(* CODESYS project DemoLib.library
   Title: DemoLib
   Author: TwinCAT Explorer
   Company: Demo
   Version: 1.0.0.0
   Placeholder: DemoLib

Project tree, tasks and I/O mapping:
  libraries: Tc2_Standard, * (Beckhoff Automation GmbH); Tc2_System, * (Beckhoff Automation GmbH)
  DUTs/
    data type E_ValveState
    data type ST_ValveStatus
    data type T_Percent
    data type U_Word
  GVLs/
    global variables GVL_DemoLib
  POUs/
    Valves/
      function block FB_ValveBase [ST]: Close, Open, State
      interface I_Valve: Close, Open, State
    function F_Clamp [ST]
  VISUs/
*)

// DUTs/E_ValveState
{attribute 'qualified_only'}
{attribute 'strict'}
TYPE E_ValveState :
(
	Closed := 0,
	Opening,
	Open,
	Closing,
	Error := 99
);
END_TYPE

// DUTs/ST_ValveStatus
TYPE ST_ValveStatus :
STRUCT
	eState		: E_ValveState;
	bInterlocked	: BOOL;
	nCycles		: UDINT;
	fOpenTime	: LREAL; // s
END_STRUCT
END_TYPE

// DUTs/T_Percent
TYPE T_Percent : LREAL;
END_TYPE

// DUTs/U_Word
TYPE U_Word :
UNION
	nValue	: WORD;
	aBytes	: ARRAY[0..1] OF BYTE;
END_UNION
END_TYPE

// GVLs/GVL_DemoLib
{attribute 'qualified_only'}
VAR_GLOBAL CONSTANT
	MAX_VALVES		: INT := 8;
	DEFAULT_TIMEOUT	: TIME := T#5S;
END_VAR

// POUs/Valves/FB_ValveBase
FUNCTION_BLOCK ABSTRACT FB_ValveBase IMPLEMENTS I_Valve
VAR_INPUT
	bInterlock	: BOOL;
END_VAR
VAR_OUTPUT
	stStatus	: ST_ValveStatus;
END_VAR
VAR
	tonTimeout	: TON;
END_VAR

tonTimeout(IN := stStatus.eState = E_ValveState.Opening OR stStatus.eState = E_ValveState.Closing, PT := GVL_DemoLib.DEFAULT_TIMEOUT);
IF tonTimeout.Q THEN
	stStatus.eState := E_ValveState.Error;
END_IF
stStatus.bInterlocked := bInterlock;

METHOD Close : BOOL
stStatus.eState := E_ValveState.Closing;
Close := TRUE;
END_METHOD

METHOD Open : BOOL
VAR_INPUT
	bForce	: BOOL;
END_VAR
IF bInterlock AND NOT bForce THEN
	RETURN;
END_IF
stStatus.eState := E_ValveState.Opening;
stStatus.nCycles := stStatus.nCycles + 1;
Open := TRUE;
END_METHOD

PROPERTY State : E_ValveState
GET
PUBLIC
VAR
END_VAR
State := stStatus.eState;
END_GET
END_PROPERTY

END_FUNCTION_BLOCK

// POUs/Valves/I_Valve
INTERFACE I_Valve

METHOD Close : BOOL
END_METHOD

METHOD Open : BOOL
VAR_INPUT
	bForce	: BOOL;
END_VAR
END_METHOD

PROPERTY State : E_ValveState
GET
PUBLIC
VAR
END_VAR
END_GET
END_PROPERTY

END_INTERFACE

// POUs/F_Clamp
FUNCTION F_Clamp : LREAL
VAR_INPUT
	fValue	: LREAL;
	fMin	: LREAL;
	fMax	: LREAL;
END_VAR

F_Clamp := MIN(MAX(fValue, fMin), fMax);

END_FUNCTION
